TYPE "st_Io_Ph_AnalogInputs"
VERSION : 0.1
   STRUCT
      Zone1_Pt1 { ExternalAccessible := 'False'; ExternalVisible := 'False'; ExternalWritable := 'False'; S7_SetPoint := 'False'} : "st_Io_Ph_AnalogInput";
      Zone1_Vacuummeter1 { ExternalAccessible := 'False'; ExternalVisible := 'False'; ExternalWritable := 'False'; S7_SetPoint := 'False'} : "st_Io_Ph_AnalogInput";
      Zone1_WaterTemperature { ExternalAccessible := 'False'; ExternalVisible := 'False'; ExternalWritable := 'False'; S7_SetPoint := 'False'} : "st_Io_Ph_AnalogInput";
      Zone1_AmbientTemperature { ExternalAccessible := 'False'; ExternalVisible := 'False'; ExternalWritable := 'False'; S7_SetPoint := 'False'} : "st_Io_Ph_AnalogInput";
      Zone1_Vibration { ExternalAccessible := 'False'; ExternalVisible := 'False'; ExternalWritable := 'False'; S7_SetPoint := 'False'} : "st_Io_Ph_AnalogInput";
      Zone1_Temperature { ExternalAccessible := 'False'; ExternalVisible := 'False'; ExternalWritable := 'False'; S7_SetPoint := 'False'} : "st_Io_Ph_AnalogInput";
      Zone1_Sound { ExternalAccessible := 'False'; ExternalVisible := 'False'; ExternalWritable := 'False'; S7_SetPoint := 'False'} : "st_Io_Ph_AnalogInput";
      Zone1_Speed { ExternalAccessible := 'False'; ExternalVisible := 'False'; ExternalWritable := 'False'; S7_SetPoint := 'False'} : "st_Io_Ph_AnalogInput";
      Zone1_Torque { ExternalAccessible := 'False'; ExternalVisible := 'False'; ExternalWritable := 'False'; S7_SetPoint := 'False'} : "st_Io_Ph_AnalogInput";
      Zone2_Pt1 { ExternalAccessible := 'False'; ExternalVisible := 'False'; ExternalWritable := 'False'; S7_SetPoint := 'False'} : "st_Io_Ph_AnalogInput";
      Zone2_Pt2 { ExternalAccessible := 'False'; ExternalVisible := 'False'; ExternalWritable := 'False'; S7_SetPoint := 'False'} : "st_Io_Ph_AnalogInput";
      Zone2_Vacuummeter1 { ExternalAccessible := 'False'; ExternalVisible := 'False'; ExternalWritable := 'False'; S7_SetPoint := 'False'} : "st_Io_Ph_AnalogInput";
      Zone2_Vacuummeter2 { ExternalAccessible := 'False'; ExternalVisible := 'False'; ExternalWritable := 'False'; S7_SetPoint := 'False'} : "st_Io_Ph_AnalogInput";
      Zone2_WaterTemperature { ExternalAccessible := 'False'; ExternalVisible := 'False'; ExternalWritable := 'False'; S7_SetPoint := 'False'} : "st_Io_Ph_AnalogInput";
      Zone2_AmbientTemperature { ExternalAccessible := 'False'; ExternalVisible := 'False'; ExternalWritable := 'False'; S7_SetPoint := 'False'} : "st_Io_Ph_AnalogInput";
      Zone2_Vibration { ExternalAccessible := 'False'; ExternalVisible := 'False'; ExternalWritable := 'False'; S7_SetPoint := 'False'} : "st_Io_Ph_AnalogInput";
      Zone2_Temperature { ExternalAccessible := 'False'; ExternalVisible := 'False'; ExternalWritable := 'False'; S7_SetPoint := 'False'} : "st_Io_Ph_AnalogInput";
      Zone2_Sound { ExternalAccessible := 'False'; ExternalVisible := 'False'; ExternalWritable := 'False'; S7_SetPoint := 'False'} : "st_Io_Ph_AnalogInput";
      Zone2_Speed { ExternalAccessible := 'False'; ExternalVisible := 'False'; ExternalWritable := 'False'; S7_SetPoint := 'False'} : "st_Io_Ph_AnalogInput";
      Zone2_Torque { ExternalAccessible := 'False'; ExternalVisible := 'False'; ExternalWritable := 'False'; S7_SetPoint := 'False'} : "st_Io_Ph_AnalogInput";
      Zone3_Pt1 { ExternalAccessible := 'False'; ExternalVisible := 'False'; ExternalWritable := 'False'; S7_SetPoint := 'False'} : "st_Io_Ph_AnalogInput";
      Zone3_Pt2 { ExternalAccessible := 'False'; ExternalVisible := 'False'; ExternalWritable := 'False'; S7_SetPoint := 'False'} : "st_Io_Ph_AnalogInput";
      Zone3_Vacuummeter1 { ExternalAccessible := 'False'; ExternalVisible := 'False'; ExternalWritable := 'False'; S7_SetPoint := 'False'} : "st_Io_Ph_AnalogInput";
      Zone3_Vacuummeter2 { ExternalAccessible := 'False'; ExternalVisible := 'False'; ExternalWritable := 'False'; S7_SetPoint := 'False'} : "st_Io_Ph_AnalogInput";
      Zone3_WaterTemperature { ExternalAccessible := 'False'; ExternalVisible := 'False'; ExternalWritable := 'False'; S7_SetPoint := 'False'} : "st_Io_Ph_AnalogInput";
      Zone3_AmbientTemperature { ExternalAccessible := 'False'; ExternalVisible := 'False'; ExternalWritable := 'False'; S7_SetPoint := 'False'} : "st_Io_Ph_AnalogInput";
      Zone3_Vibration { ExternalAccessible := 'False'; ExternalVisible := 'False'; ExternalWritable := 'False'; S7_SetPoint := 'False'} : "st_Io_Ph_AnalogInput";
      Zone3_Temperature { ExternalAccessible := 'False'; ExternalVisible := 'False'; ExternalWritable := 'False'; S7_SetPoint := 'False'} : "st_Io_Ph_AnalogInput";
      Zone3_Sound { ExternalAccessible := 'False'; ExternalVisible := 'False'; ExternalWritable := 'False'; S7_SetPoint := 'False'} : "st_Io_Ph_AnalogInput";
      Zone3_Speed { ExternalAccessible := 'False'; ExternalVisible := 'False'; ExternalWritable := 'False'; S7_SetPoint := 'False'} : "st_Io_Ph_AnalogInput";
      Zone3_Torque { ExternalAccessible := 'False'; ExternalVisible := 'False'; ExternalWritable := 'False'; S7_SetPoint := 'False'} : "st_Io_Ph_AnalogInput";
      Zone1_FM1 { ExternalAccessible := 'False'; ExternalVisible := 'False'; ExternalWritable := 'False'; S7_SetPoint := 'False'} : "st_Io_Ph_AnalogInput";
      Zone1_FM2 { ExternalAccessible := 'False'; ExternalVisible := 'False'; ExternalWritable := 'False'; S7_SetPoint := 'False'} : "st_Io_Ph_AnalogInput";
      Zone2_FM1 { ExternalAccessible := 'False'; ExternalVisible := 'False'; ExternalWritable := 'False'; S7_SetPoint := 'False'} : "st_Io_Ph_AnalogInput";
      Zone2_FM2 { ExternalAccessible := 'False'; ExternalVisible := 'False'; ExternalWritable := 'False'; S7_SetPoint := 'False'} : "st_Io_Ph_AnalogInput";
      Zone2_FM3 { ExternalAccessible := 'False'; ExternalVisible := 'False'; ExternalWritable := 'False'; S7_SetPoint := 'False'} : "st_Io_Ph_AnalogInput";
      Zone2_FM4 { ExternalAccessible := 'False'; ExternalVisible := 'False'; ExternalWritable := 'False'; S7_SetPoint := 'False'} : "st_Io_Ph_AnalogInput";
      Zone3_FM1 { ExternalAccessible := 'False'; ExternalVisible := 'False'; ExternalWritable := 'False'; S7_SetPoint := 'False'} : "st_Io_Ph_AnalogInput";
      Zone3_FM2 { ExternalAccessible := 'False'; ExternalVisible := 'False'; ExternalWritable := 'False'; S7_SetPoint := 'False'} : "st_Io_Ph_AnalogInput";
      Zone3_FM3 { ExternalAccessible := 'False'; ExternalVisible := 'False'; ExternalWritable := 'False'; S7_SetPoint := 'False'} : "st_Io_Ph_AnalogInput";
      Zone3_FM4 { ExternalAccessible := 'False'; ExternalVisible := 'False'; ExternalWritable := 'False'; S7_SetPoint := 'False'} : "st_Io_Ph_AnalogInput";
   END_STRUCT;

END_TYPE

